// TIA Portal V21 export
ORGANIZATION_BLOCK "Timer"   // OB1, LAD
BEGIN

REGION Network 1: Start delay
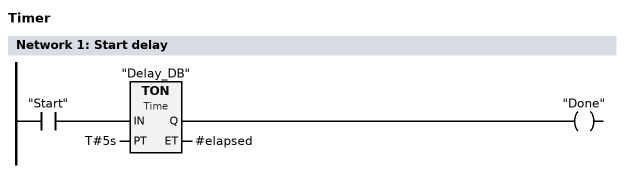
   RUNG wire#powerrail
      Contact( "Start" )
      { S7_Templates := "time_type := Time" } "Delay_DB".TON(pt := T#5s, et => #elapsed)
      Coil( "Done" )
   END_RUNG
   // the same network as SCL:
   "Delay_DB".TON(IN := "Start", PT := T#5s, ET => #elapsed);
   "Done" := "Delay_DB".Q;
END_REGION
END_ORGANIZATION_BLOCK
